// TIA Portal V21 export
// export: Created 2026-11-11T00:47:21.239823Z, ExportSetting WithDefaults, DisplayName Totally Integrated Automation Portal, DisplayVersion V21 Update 3, DisplayName STEP 7 Professional, DisplayVersion V21 Update 3, DisplayName STEP 7 Safety, DisplayVersion V21, DisplayName Tech WebApplication, DisplayVersion V21, DisplayName WinCC Basic/Comfort/Advanced, DisplayVersion V21 Update 3, DisplayName WinCC Unified, DisplayVersion V21 Update 3
FUNCTION_BLOCK "FB_Fbd_ex062"   // FB98, FBD
{ S7_Optimized_Access := 'TRUE' }
VERSION : 0.1
// stored: AutoNumber true, IsIECCheckEnabled false, IsRetainMemResEnabled false, MemoryReserve 100, SetENOAutomatically false, UDAEnableTagReadback false
   VAR_INPUT
      v_mode : Int;
      v_f_id : HW_SUBMODULE;
      v_mlen : Int;
      v_code1 : Byte;
      v_code2 : Byte;
   END_VAR
   VAR_OUTPUT
      v_new : Bool;
      v_status : DWord;
      v_slot : HW_SUBMODULE;
      v_subslot : HW_SUBMODULE;
      v_index : UInt;
      v_len : UInt;
   END_VAR
   VAR_IN_OUT
      v_record : Array[0..99] of Byte;
   END_VAR
   VAR
      inst { S7_SetPoint := 'True'} : RCVREC;
   END_VAR
BEGIN

REGION Network 1: RCVREC - Receive data record
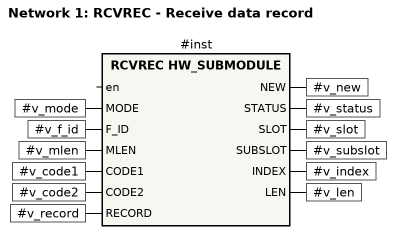
   #inst(MODE := #v_mode,   // RCVREC
         F_ID := #v_f_id,
         MLEN := #v_mlen,
         CODE1 := #v_code1,
         CODE2 := #v_code2,
         RECORD := #v_record,
         NEW => #v_new,
         STATUS => #v_status,
         SLOT => #v_slot,
         SUBSLOT => #v_subslot,
         INDEX => #v_index,
         LEN => #v_len);
END_REGION
END_FUNCTION_BLOCK
